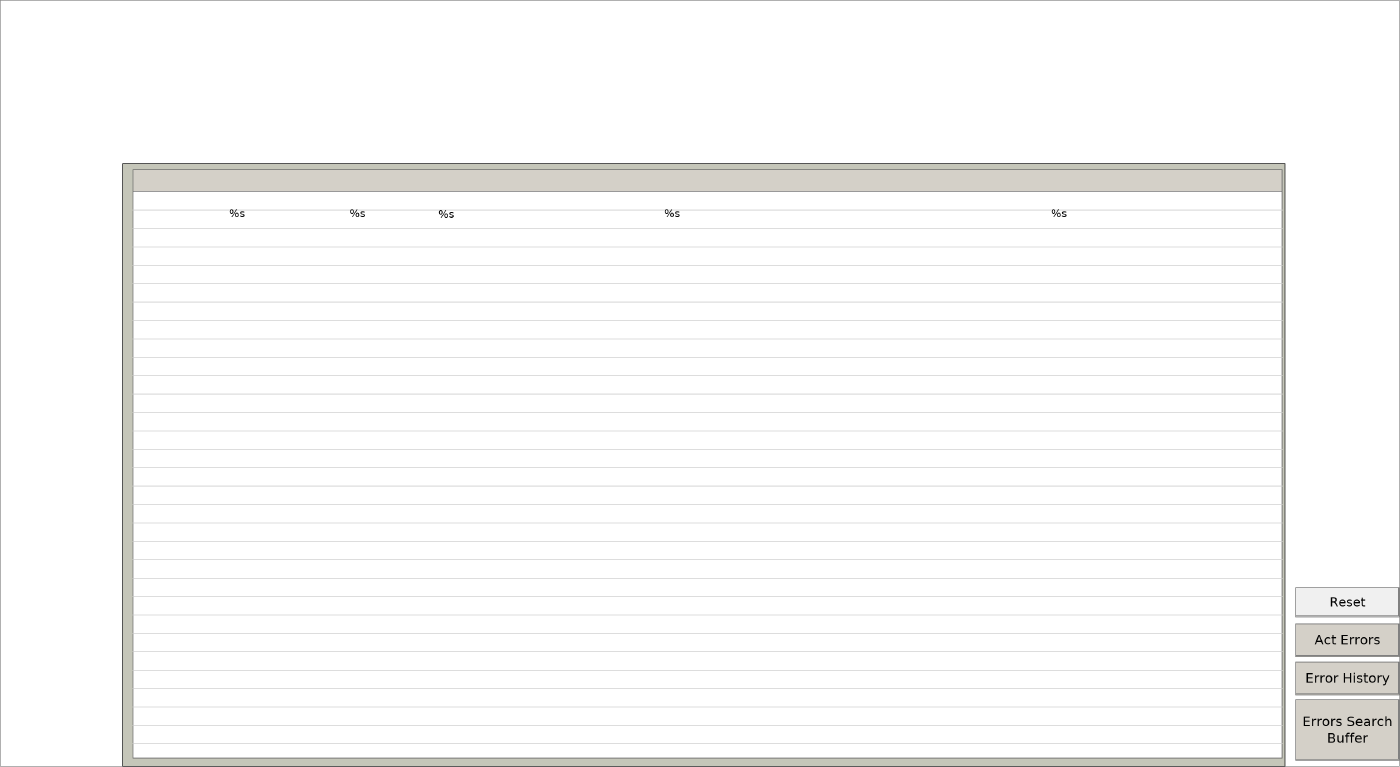
VISUALIZATION ERROR_BUFFER  // 1900x1042
    Group (1758,798 142x235)
        Button (0,0 142x40), "Reset", pressed state: prg_Messages.ResetErrors
            toggle prg_Messages.ResetErrors
        Button (0,101 142x45), "Error History"
            OnMouseClick: change screen: ERROR_HISTORY
        Button (0,152 142x83), "Errors Search Buffer"
            OnMouseClick: change screen: ERROR_BUFFER
        Button (0,49 142x45), "Act Errors"
            OnMouseClick: change screen: ERRORS_OPER
    Rectangle (166,222 1578x820)
    Table (180,230 1560x800), data array: Buffer_Search_Messages
        p3854506369: Buffer_Search_Messages[INDEX].sDateTime
        p1892666644: Buffer_Search_Messages[INDEX].sErrID
        p338671338: Buffer_Search_Messages[INDEX].sLevel
        p2170511999: Buffer_Search_Messages[INDEX].sModuleDescription
        p3723444502: Buffer_Search_Messages[INDEX].sErrorMessage
        p4092479075: Module Description
        p2237128397: Error Message
    Rectangle (421,270 129x40), "%s", text variable: Prg_Filter_Messages.stFilter.sErrID
        OnMouseClick: write the text variable via Edit
    Rectangle (551,271 110x40), "%s", text variable: Prg_Filter_Messages.stFilter.sLevel
        OnMouseClick: write the text variable via Edit
    Rectangle (662,270 501x40), "%s", text variable: Prg_Filter_Messages.stFilter.sModuleDescription
        OnMouseClick: write the text variable via Edit
    Rectangle (1162,270 551x40), "%s", text variable: Prg_Filter_Messages.stFilter.sErrorMessage
        OnMouseClick: write the text variable via Edit
    Rectangle (222,270 200x40), "%s", text variable: Prg_Filter_Messages.stFilter.sDateTime
        OnMouseClick: write the text variable via Edit
END_VISUALIZATION

(* stored: Version 1.1.0.1, ProductVersion 3.1.4024.13
   Visu ERROR_BUFFER: Id {714473b8-d707-4ec7-8870-c8afe1d19a50} *)
